FUNCTION_BLOCK Valvula_Solenoide (* Valvula solenoide on/off (saida digital) com fim de curso opcional - HidrycoLib *)
  (* Standard: 61499-2 *)
  (* Version 1.0, 04/11/2026, Hidryco, Hidryco, 1.0: SV-900 da agua de servico do lodo. O comando continua na logica do pai (cmdAbrir com REQ). Fins de curso por symlink ${PATH}stsAberto e ${PATH}stsFechado, usados so com cfgUsaFimCurso = TRUE; sem eles aberta/fechada saem do comando. Alarme = discrepancia por cfgTempoFalha (s). Modo sempre manual (fbkStsAutomatico = FALSE). *)
  PACKAGE Hidryco.HidrycoLib;
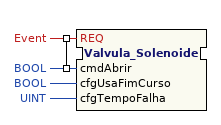
  EVENT_INPUT
    REQ WITH cmdAbrir; (* Novo comando da logica *)
  END_EVENT
  VAR_INPUT
    cmdAbrir : BOOL; (* Comando abrir (mesmo valor enviado a saida digital) *)
    cfgUsaFimCurso : BOOL := FALSE; (* TRUE = usa os fins de curso (symlinks stsAberto/stsFechado) e alarme de discrepancia *)
    cfgTempoFalha : UINT := 10; (* Tempo de discrepancia para o alarme (s) *)
  END_VAR
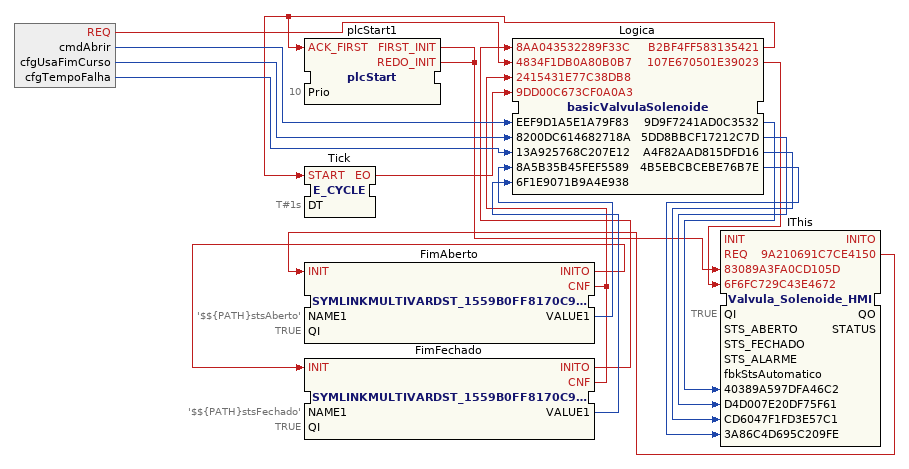
  FBS
    IThis : Valvula_Solenoide_HMI(QI := TRUE);
    plcStart1 : plcStart(Prio := 10);
    Tick : E_CYCLE(DT := T#1s);
    Logica : basicValvulaSolenoide;
    FimAberto : SYMLINKMULTIVARDST_1559B0FF8170C9BA0(NAME1 := '$${PATH}stsAberto', QI := TRUE); {SET_ATTRIBUTE(Configuration.GenericFBType.InterfaceParams, Runtime.System#I:=1;VALUE${I$}:BOOL)}
    FimFechado : SYMLINKMULTIVARDST_1559B0FF8170C9BA0(NAME1 := '$${PATH}stsFechado', QI := TRUE); {SET_ATTRIBUTE(Configuration.GenericFBType.InterfaceParams, Runtime.System#I:=1;VALUE${I$}:BOOL)}
  END_FBS
  EVENT_CONNECTIONS
    plcStart1.FIRST_INIT TO IThis.83089A3FA0CD105D;
    plcStart1.REDO_INIT TO IThis.83089A3FA0CD105D;
    IThis.9A210691C7CE4150 TO FimAberto.INIT;
    FimAberto.INITO TO FimFechado.INIT;
    FimFechado.INITO TO Logica.8AA043532289F33C;
    Logica.B2BF4FF583135421 TO Tick.START;
    Logica.B2BF4FF583135421 TO plcStart1.ACK_FIRST;
    REQ TO Logica.4834F1DB0A80B0B7;
    FimAberto.CNF TO Logica.2415431E77C38DB8;
    FimFechado.CNF TO Logica.2415431E77C38DB8;
    Tick.EO TO Logica.9DD00C673CF0A0A3;
    Logica.107E670501E39023 TO IThis.6F6FC729C43E4672;
  END_CONNECTIONS
  DATA_CONNECTIONS
    cmdAbrir TO Logica.EEF9D1A5E1A79F83;
    cfgUsaFimCurso TO Logica.8200DC614682718A;
    cfgTempoFalha TO Logica.13A925768C207E12;
    FimAberto.VALUE1 TO Logica.8A5B35B45FEF5589;
    FimFechado.VALUE1 TO Logica.6F1E9071B9A4E938;
    Logica.9D9F7241AD0C3532 TO IThis.40389A597DFA46C2;
    Logica.5DD8BBCF17212C7D TO IThis.D4D007E20DF75F61;
    Logica.A4F82AAD815DFD16 TO IThis.CD6047F1FD3E57C1;
    Logica.4B5EBCBCEBE76B7E TO IThis.3A86C4D695C209FE;
  END_CONNECTIONS
END_FUNCTION_BLOCK
